# EPICS substitutions: db/Beckhoff_7XXX/ecmcEX72XX_OPT_info2Temp.substitutions
file "ecmc_analogInput-chX.template"
{
  pattern {CH_ID, sourceName, KEY, suffix, DESC, EGU, ESLO, PREC, LOPR, HOPR, LOLO, LOW, HIGH, HIHI, HYST, LLSV, LSV, HSV, HHSV}
          {"$(OPT_CH_ID=01)", "temperatureActual", "Drv", "-TmpAct", "PCB temperature", "degC", 0.1, 1, 0, 50, 0, 0, 40, 50, 0.5, "NO_ALARM", "NO_ALARM", "MINOR", "MAJOR"}
}
